FUNCTION_BLOCK abs_a
VAR_INPUT
	x: ARRAY[0..243] OF LREAL;
END_VAR
VAR_OUTPUT
	y: ARRAY[0..243] OF LREAL;
END_VAR
VAR
	k: DINT;
END_VAR



FOR k := 0 TO 243 DO 
    y[k] := ABS(x[k]);
END_FOR;

END_FUNCTION_BLOCK

(* stored: Version 1.1.0.1, ProductVersion 3.1.4024.9
   POU abs_a: Id {dde1d8f0-9800-4053-b040-44a116a490ae}, SpecialFunc None *)
